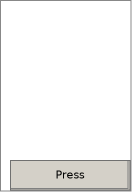
VISUALIZATION VisuE4x  // 132x192
    Button (10,160 120x30), "Press", pressed state: GVL_Fixture.bEnable
END_VISUALIZATION

(* stored: Version 1.1.0.1
   Visu VisuE4x: Id {67b51daa-a272-43b9-8df9-e19dc83959c5} *)
